(* IEC 61131-3 sources: Test-Git_ESME26/TestProgettoESME_26.fbsproj/AxisModuleLib Migration, 10 files *)

(* ---- AXM_GPL.gvl ---- *)
{attribute 'qualified_only'}
VAR_GLOBAL CONSTANT
	Gc_udiMaxNumberOfCamTables		: UDINT := 4;
END_VAR

(* ---- AXM_FC_EtCmdToString.fn.st ---- *)
FUNCTION PUBLIC AXM_FC_EtCmdToString : STRING[20]
VAR_INPUT
	i_etCmd : AXM_ET_Cmd;
END_VAR
VAR_OUTPUT
	q_etDiag	: GD.ET_Diag := GD.ET_Diag.Ok;
	q_etDiagExt	: AXM_ET_DiagExt := AXM_ET_DiagExt.Ok;
END_VAR
VAR
END_VAR

AXM_FC_EtCmdToString := TO_STRING(i_etCmd);
IF TO_UDINT(AXM_FC_EtCmdToString) <> 0 THEN // if the string is not a number the result is 0
	AXM_FC_EtCmdToString := Standard.CONCAT('Unknown DiagExt: ', TO_STRING(i_etCmd));
	q_etDiag := GD.ET_Diag.InputParameterInvalid;
	q_etDiagExt := AXM_ET_DiagExt.CmdUnknown;;
END_IF

(* ---- AXM_FC_EtMotionActiveVelTypeToString.fn.st ---- *)
FUNCTION PUBLIC AXM_FC_EtMotionActiveVelTypeToString : STRING[20]
VAR_INPUT
	i_etMotionActiveVelType : AXM_ET_MotionActiveVelType;
END_VAR
VAR_OUTPUT
	q_etDiag	: GD.ET_Diag := GD.ET_Diag.Ok;
	q_etDiagExt	: AXM_ET_DiagExt := AXM_ET_DiagExt.Ok;
END_VAR
VAR
END_VAR

AXM_FC_EtMotionActiveVelTypeToString := TO_STRING(i_etMotionActiveVelType);

(* ---- AXM_FC_EtOpModeToString.fn.st ---- *)
FUNCTION PUBLIC AXM_FC_EtOpModeToString : STRING[20]
VAR_INPUT
	i_etOpMode : AXM_ET_OpMode;
END_VAR
VAR_OUTPUT
	q_etDiag	: GD.ET_Diag := GD.ET_Diag.Ok;
	q_etDiagExt	: AXM_ET_DiagExt := AXM_ET_DiagExt.Ok;
END_VAR
VAR
END_VAR

AXM_FC_EtOpModeToString := TO_STRING(i_etOpMode);

(* ---- AXM_FC_EtParIdToString.fn.st ---- *)
FUNCTION PUBLIC AXM_FC_EtParIdToString : STRING[20]
VAR_INPUT
	i_etParId : AXM_ET_ParId;
END_VAR
VAR_OUTPUT
	q_etDiag	: GD.ET_Diag := GD.ET_Diag.Ok;
	q_etDiagExt	: AXM_ET_DiagExt := AXM_ET_DiagExt.Ok;
END_VAR
VAR
END_VAR

AXM_FC_EtParIdToString := TO_STRING(i_etParId);

(* ---- AXM_FC_EtStateToString.fn.st ---- *)
FUNCTION PUBLIC AXM_FC_EtStateToString : String[80]
VAR_INPUT
	i_etState	: AXM_ET_State;
END_VAR
VAR_OUTPUT
	q_etDiag	: GD.ET_Diag := GD.ET_Diag.Ok;
	q_etDiagExt	: AXM_ET_DiagExt := AXM_ET_DiagExt.Ok;
END_VAR
VAR
END_VAR

AXM_FC_EtStateToString := TO_STRING(i_etState);

(* ---- AXM_FC_UpdateAddInterfaceStruct.fn.st ---- *)
/// FC version: 1.0.0.0
/// Example Project version: 26.0.11.0 (Automatically generated, do not change!)

FUNCTION PUBLIC AXM_FC_UpdateAddInterfaceStruct : BOOL
VAR_INPUT
	i_pdwSubModuleAddInterfaces : POINTER TO TPL.TYPE_ADDRESS; // change from DWORD to TYPE_ADDRESS;
	i_udiSubModuleConstant		: UDINT;
END_VAR
VAR_IN_OUT
	iq_stAxisModuleItf	: AXM_ST_ModuleInterface;
END_VAR
VAR_OUTPUT
	q_etDiag			: GD.ET_Diag := GD.ET_Diag.Ok;
	q_etDiagExt			: AXM_ET_DiagExt := AXM_ET_DiagExt.Ok;
	q_sMsg				: STRING[80];
END_VAR
VAR
	pdwArrayPos			: POINTER TO TPL.TYPE_ADDRESS; // change from DWORD to TYPE_ADDRESS;
END_VAR

(********************************************************************************************************
revision history:
=========================================================================================================
version	|	date		| author				| comment
=========================================================================================================
1.0.0.0	|	2025-03-18	| Schneider Electric	| - initial release
---------------------------------------------------------------------------------------------------------
1.x.y.z	|	20xx-xx-xx	| your name				| - What has been modified?
=========================================================================================================
********************************************************************************************************)

IF i_pdwSubModuleAddInterfaces = 0 THEN
	q_etDiag	:= GD.ET_Diag.InputParameterInvalid;
	q_etDiagExt	:= AXM_ET_DiagExt.SubModuleAddInterfacesInvalidPointer;
	q_sMsg		:= '';
ELSIF i_udiSubModuleConstant < 1 THEN
	q_etDiag	:= GD.ET_Diag.InputParameterInvalid;
	q_etDiagExt := AXM_ET_DiagExt.SubModuleConstantRange;
	q_sMsg		:= '1 <= i_udiSubModuleConstant';
ELSE
	pdwArrayPos := i_pdwSubModuleAddInterfaces + (i_udiSubModuleConstant-1) * SIZEOF(pdwArrayPos^);
	pdwArrayPos^ := ADR(iq_stAxisModuleItf);
END_IF

(* ---- AXM_FB_AxisModuleController.fb.st ---- *)
FUNCTION_BLOCK PUBLIC AXM_FB_AxisModuleController
VAR_INPUT
	i_xEnable			: BOOL;
END_VAR
VAR_IN_OUT
	iq_stStandardModuleItf			: TPL.ST_StandardModuleInterface;
	iq_stStandardMotionItf			: TPL.ST_StandardMotionInterface;
	iq_stExceptionList				: TPL.ST_ExceptionList;
	iq_stLogDataList				: TPL.ST_LogDataList;
END_VAR
VAR_OUTPUT
	q_xActive			: BOOL;
	q_xReady			: BOOL;
	q_etDiag			: GD.ET_Diag := GD.ET_Diag.Ok;
	q_etDiagExt			: AXM_ET_DiagExt := AXM_ET_DiagExt.Disabled;
	q_sMsg				: STRING[80] := '';
END_VAR
VAR
	pdw								: POINTER TO TPL.TYPE_ADDRESS; // change from DWORD to TYPE_ADDRESS;
	udiModul						: UDINT;
	pstStandardInterface			: POINTER TO TPL.ST_StandardModuleInterface;
	pstAxisInterface				: POINTER TO AXM_ST_ModuleInterface;
	xSercState						: BOOL;
	xSercStateOld					: BOOL := TRUE;
	xJogForwEdgeDetect              : BOOL := FALSE;
	xJogBackEdgeDetect              : BOOL := FALSE;
END_VAR

IF i_xEnable AND NOT q_xActive THEN
	q_xActive := TRUE;
	q_xReady := TRUE;
	q_etDiag := GD.ET_Diag.Ok;
	q_etDiagExt := AXM_ET_DiagExt.Working;
	q_sMsg		:= '';
ELSIF NOT i_xEnable AND q_xActive THEN
	IF(iq_stStandardModuleItf.iq_stExt.dwSubModulesItf <> 0 AND iq_stStandardModuleItf.iq_stExt.pdwSubModulesAddItf <> 0) THEN
		FOR udiModul:= 1 TO iq_stStandardModuleItf.iq_stExt.udiNumberOfSubModules DO
			pstStandardInterface := iq_stStandardModuleItf.iq_stExt.dwSubModulesItf + UDINT_TO_DWORD((udiModul - 1) * SIZEOF(pstStandardInterface^));
			IF(pstStandardInterface^.q_dwModuleType = UDINT_TO_DWORD(TPL.ET_ModuleType.AxisModule)) THEN
				(* Module version check *)
				IF(pstStandardInterface^.q_udiModuleVersion = 1) THEN
					pdw := iq_stStandardModuleItf.iq_stExt.pdwSubModulesAddItf + UDINT_TO_DWORD((udiModul - 1) * SIZEOF(pdw^));
					pstAxisInterface := pdw^;
					IF(pstAxisInterface <> 0) THEN
						pstAxisInterface^.stManual.i_xJogForw := FALSE;
						pstAxisInterface^.stManual.i_xJogBack := FALSE;
					END_IF
				END_IF
			END_IF
		END_FOR
	END_IF
	q_xReady 	:= FALSE;
	q_xActive	:= FALSE;
	q_etDiag	:= GD.ET_Diag.Ok;
	q_etDiagExt	:= AXM_ET_DiagExt.Disabled;
	q_sMsg		:= '';
END_IF
IF ((iq_stStandardModuleItf.iq_stExt.udiNumberOfSubModules <> 0)
	AND ((iq_stStandardModuleItf.iq_stExt.pdwSubModulesAddItf = 0) OR (iq_stStandardModuleItf.iq_stExt.dwSubModulesItf = 0))) THEN
	q_xReady := FALSE;
	q_etDiag := GD.ET_Diag.InputParameterInvalid;
	q_etDiagExt := AXM_ET_DiagExt.MissingExtInit;
	q_sMsg := 'Missing Call of FC_UpdateAddInterfaceStruct';
END_IF

IF q_xActive AND q_xReady  THEN
 	IF (FC_GetSercosState() >= SMI.ET_SercosState.NRT) THEN
		xSercState := (FC_GetSercosState() = SMI.ET_SercosState.Phase4);
		IF(iq_stStandardModuleItf.iq_stExt.dwSubModulesItf <> 0 AND iq_stStandardModuleItf.iq_stExt.pdwSubModulesAddItf <> 0) THEN
			FOR udiModul := 1 TO iq_stStandardModuleItf.iq_stExt.udiNumberOfSubModules DO
				pstStandardInterface := iq_stStandardModuleItf.iq_stExt.dwSubModulesItf + UDINT_TO_DWORD((udiModul - 1) * SIZEOF(pstStandardInterface^));
				IF(pstStandardInterface^.q_dwModuleType = TPL.ET_ModuleType.AxisModule) THEN
					(* Module version check *)
					IF(pstStandardInterface^.q_udiModuleVersion = 1) THEN
						pdw := iq_stStandardModuleItf.iq_stExt.pdwSubModulesAddItf +  UDINT_TO_DWORD((udiModul - 1) * SIZEOF(pdw^));
						IF(pdw^ = 0) THEN (* Configuration error in stSubModules *)
							q_xReady := FALSE;
							q_etDiag := GD.ET_Diag.InputParameterInvalid;
							q_etDiagExt := AXM_ET_DiagExt.MissingExtInit;
							q_sMsg := 'Missing Call of FC_UpdateAddInterfaceStruct';
							RETURN;
						END_IF
						pstAxisInterface := pdw^;
						IF(pstAxisInterface <> 0) THEN
							(* Implementation of axis select *)
							IF iq_stStandardMotionItf.i_udiModuleSelect > 0 AND iq_stStandardMotionItf.i_udiModuleSelect = pstStandardInterface^.i_udiModuleId THEN

								(* Don't set pstAxisInterface^.stManual.i_xJog* from iq_stStandardMotionItf.i_xJog* blindly since the Vis might want to jog as well *)
								IF (iq_stStandardMotionItf.i_xJogForw) THEN
									pstAxisInterface^.stManual.i_xJogForw := TRUE;
									xJogForwEdgeDetect := TRUE;
								ELSE
									IF (xJogForwEdgeDetect) THEN
										pstAxisInterface^.stManual.i_xJogForw := FALSE;
										xJogForwEdgeDetect := FALSE;
								    END_IF
								END_IF
								IF (iq_stStandardMotionItf.i_xJogBack) THEN
									pstAxisInterface^.stManual.i_xJogBack := TRUE;
									xJogBackEdgeDetect := TRUE;
								ELSE
									IF (xJogBackEdgeDetect) THEN
										pstAxisInterface^.stManual.i_xJogBack := FALSE;
										xJogBackEdgeDetect := FALSE;
								    END_IF
								END_IF

							ELSE
								pstAxisInterface^.stManual.i_xJogForw := FALSE;
								pstAxisInterface^.stManual.i_xJogBack := FALSE;
							END_IF
							(* Implementation of HomeOkReset *)
							IF NOT xSercState  THEN (* As long as the sercos state is <> 4, set the reset home ok to true *)
								pstAxisInterface^.stHome.i_xResetHomeOk := TRUE;
							ELSIF NOT xSercStateOld THEN (* Detect a positive edge in xSercState, the sercos has entered state 4 *)
								pstAxisInterface^.stHome.i_xResetHomeOk := FALSE;
							END_IF
						END_IF
					END_IF
				END_IF
			END_FOR
 		END_IF
	ELSE
		xSercState := FALSE;
		q_xReady := FALSE;
		q_etDiag := GD.ET_Diag.SercosConditionInvalid;
		q_etDiagExt := AXM_ET_DiagExt.GlobalSercosInterfaceInvalid;
		q_sMsg := AXM_FC_EtDiagExtToString(i_etDiagExt := AXM_ET_DiagExt.GlobalSercosInterfaceInvalid);
	END_IF
	xSercStateOld := xSercState;
END_IF

(* ---- AXM_FB_AxisModuleVisController.fb.st ---- *)
FUNCTION_BLOCK PUBLIC AXM_FB_AxisModuleVisController
VAR_INPUT
	i_xEnable               : BOOL;
	i_pstMachineStandardItf : POINTER TO TPL.ST_StandardModuleInterface;
	i_pstCurrentStandardItf : POINTER TO TPL.ST_StandardModuleInterface;
	i_dwCurrentAddItf       : TPL.TYPE_ADDRESS; // change DWORD to TYPE_ADDRESS
	i_xUpdateData           : BOOL;
	i_udiCurrentJogTarget   : UDINT;
END_VAR
VAR_IN_OUT
	iq_stExceptionList : TPL.ST_ExceptionList;
	iq_stLogDataList   : TPL.ST_LogDataList;
END_VAR
VAR_OUTPUT
	q_xActive                          : BOOL;
	q_xReady                           : BOOL;
	q_etDiag                           : GD.ET_Diag := GD.ET_Diag.Ok;
	q_etDiagExt                        : AXM_ET_DiagExt := AXM_ET_DiagExt.Disabled;
	q_sMsg                             : STRING[80] := '';
	q_udiSetAsCurrentModule            : UDINT;
	q_udiSetAsJogTarget                : UDINT;
	q_xSimulateExceptionStopEndOfCycle : BOOL;
END_VAR
VAR
	xEnableFlag              : BOOL;
	pstCurrentAxisInterface  : POINTER TO AXM_ST_ModuleInterface;
	stOldAxisInterface       : AXM_ST_ModuleInterface;
	pstCurrent               : POINTER TO TPL.ST_StandardModuleInterface;
	xInitUserInputs          : BOOL;
	dwOldCurrentAddInterface : TPL.TYPE_ADDRESS; // change DWORD to TYPE_ADDRESS
	xSuccess                 : BOOL;
END_VAR
VAR
	viq_stCurrentAxisInterface      : AXM_ST_ModuleInterface;
	viq_pstCurrentStandardInterface : POINTER TO TPL.ST_StandardModuleInterface;
	vq_xCurrentIsOfMyType           : BOOL;
	vi_iPaneSelect                  : INT  := 1;
	vq_iShowOpMode                  : DINT := -1;
	vq_sOpMode                      : STRING[40];
	vi_iSelectOpMode                : INT  := -1;
	vq_sDriveName                   : STRING[40];
	vq_lrDriveRefPosition           : LREAL;
	vq_uiDriveTopologyAddress       : UINT;
	vq_diDriveState                 : DINT;
	vq_diDriveDiagCode              : DINT;
	vq_sDriveDiagMsg                : STRING[39];
	vq_lrDriveMaxVel                : LREAL;
	vq_lrDriveMaxAcc                : LREAL;
	vq_xDriveControllerEnable       : BOOL;
	vq_diDriveWorkingState          : DINT;
	vq_sMasterName                  : STRING[40];
	vq_xTpValue                     : BOOL;
	viq_xCmdStart                   : BOOL;
	viq_xCmdWSStart                 : BOOL;
	viq_xCmdHold                    : BOOL;
	viq_xDriveEnableOn              : BOOL;
	viq_xDriveEnableOff             : BOOL;
	viq_xReactionEndOfCycle         : BOOL;
	viq_xHomeLimitSwitchInvisible   : BOOL;
	viq_xHomeMoveOnPosInvisible     : BOOL;
	viq_xHomeSensorInvisible        : BOOL;
	viq_xHomeSetPosInvisible        : BOOL;
	viq_xHomeTorqueInvisible        : BOOL;
	viq_xHomeTouchProbeInvisible    : BOOL;
	viq_xHomeWritePosInvisible      : BOOL;
	viq_xHomeForceInvisible         : BOOL;
	viq_xJogForw                    : BOOL;
	viq_xJogBack                    : BOOL;
	xJogForwEdgeDetect              : BOOL := FALSE;
	xJogBackEdgeDetect              : BOOL := FALSE;
	viq_xEditCamTablesInvisible     : BOOL := TRUE;
	viq_udiEditCamTablesTableNo     : UDINT := 4;
	viq_diEditCamTablesPointNo      : DINT := 0;
	v_xHideTabHandler               : BOOL := TRUE;
	ifDiagnostic                    : UFMPLCI.IF_Diagnostic;
	ifDiagnosticAccess              : UFMPLCI.IF_DiagnosticAccess;
	ifGetParentDevice               : DTSI.IF_GetParentDevice;
	ifDeviceAccess                  : DTSI.IF_DeviceAccess;
	ifSercosIdentificationAccess    : SDI.IF_SercosIdentificationAccess;
	ifSercosIdentification          : SDI.IF_SercosIdentification;
	ifWorkingModeAccess             : CFDI.IF_WorkingModeAccess;
	ifWorkingMode                   : CFDI.IF_WorkingMode;
	ifDeviceTreeObjectSlaveAccess   : UFMPLCI.IF_DeviceTreeObjectAccess;
	ifDeviceTreeObjectMasterAccess  : UFMPLCI.IF_DeviceTreeObjectAccess;
	ifDriveConfigAccess             : DDI.IF_DriveConfigAccess;
	ifDriveConfig                   : DDI.IF_DriveConfig;
	ifOldMaster                     : MOIN.IF_Axis;
	ifTouprobeData                  : IODI.IF_TouchprobeData;
	ifTouprobeDataAccess            : IODI.IF_TouchprobeDataAccess;

END_VAR

q_udiSetAsCurrentModule            := 0;
q_udiSetAsJogTarget                := 0;
pstCurrent                         := i_pstCurrentStandardItf;
q_xSimulateExceptionStopEndOfCycle := viq_xReactionEndOfCycle;

// Calculate Homing mode invisible BOOLs
viq_xHomeLimitSwitchInvisible := viq_stCurrentAxisInterface.stHome.i_etMode < 8 OR viq_stCurrentAxisInterface.stHome.i_etMode > 11;
viq_xHomeMoveOnPosInvisible   := viq_stCurrentAxisInterface.stHome.i_etMode <> 14;
viq_xHomeSensorInvisible      := viq_stCurrentAxisInterface.stHome.i_etMode < 4 OR viq_stCurrentAxisInterface.stHome.i_etMode > 7;
viq_xHomeSetPosInvisible      := viq_stCurrentAxisInterface.stHome.i_etMode < 15 OR viq_stCurrentAxisInterface.stHome.i_etMode > 19;
viq_xHomeTorqueInvisible      := viq_stCurrentAxisInterface.stHome.i_etMode < 12 OR viq_stCurrentAxisInterface.stHome.i_etMode > 13;
viq_xHomeTouchProbeInvisible  := viq_stCurrentAxisInterface.stHome.i_etMode < 0 OR viq_stCurrentAxisInterface.stHome.i_etMode > 3;
viq_xHomeWritePosInvisible    := viq_stCurrentAxisInterface.stHome.i_etMode <> 20;
viq_xHomeForceInvisible       := viq_stCurrentAxisInterface.stHome.i_etMode < 21 OR viq_stCurrentAxisInterface.stHome.i_etMode > 22;

IF i_xEnable THEN
	q_xActive := TRUE;
	IF (i_pstCurrentStandardItf = 0) THEN
		q_xReady    := FALSE;
		q_etDiag    := GD.ET_Diag.InputParameterInvalid;
		q_etDiagExt := AXM_ET_DiagExt.CurrentStandardItfInvalid;
		q_sMsg      := 'pointer is null';
	ELSIF (i_dwCurrentAddItf = 0) THEN
		q_xReady    := FALSE;
		q_etDiag    := GD.ET_Diag.InputParameterInvalid;
		q_etDiagExt := AXM_ET_DiagExt.CurrentAddItfInvalid;
		q_sMsg      := 'pointer is null';
	ELSE
		q_xReady    := TRUE;
		q_etDiag    := GD.ET_Diag.Ok;
		q_etDiagExt := AXM_ET_DiagExt.Working;
		q_sMsg      := AXM_FC_EtDiagExtToString(i_etDiagExt := AXM_ET_DiagExt.Working);
		IF (i_pstCurrentStandardItf^.q_dwModuleType = UDINT_TO_DWORD(TPL.ET_ModuleType.AxisModule)) THEN
			(* Module version check *)
			IF (i_pstCurrentStandardItf^.q_udiModuleVersion = 1) THEN
				pstCurrentAxisInterface := i_dwCurrentAddItf;
				vq_xCurrentIsOfMyType   := TRUE;
			END_IF
		ELSE
			pstCurrentAxisInterface := 0;
			vq_xCurrentIsOfMyType   := FALSE;
		END_IF

		IF (vq_xCurrentIsOfMyType) THEN
			(* Execute changes requested by user first *)
			IF (NOT xInitUserInputs) THEN
				xInitUserInputs := TRUE;
				(* Ignore values of variables now *)
			ELSE
				DetectUserChanges();
			END_IF

			IF dwOldCurrentAddInterface <> i_dwCurrentAddItf THEN
				dwOldCurrentAddInterface        := i_dwCurrentAddItf;
				viq_stCurrentAxisInterface      := pstCurrentAxisInterface^;
				stOldAxisInterface              := viq_stCurrentAxisInterface;
				viq_pstCurrentStandardInterface := i_pstCurrentStandardItf;

				IF (viq_stCurrentAxisInterface.stMain.i_ifDrive <> 0) THEN
					xSuccess := __QUERYINTERFACE(viq_stCurrentAxisInterface.stMain.i_ifDrive, ifGetParentDevice);
					IF xSuccess THEN
						ifDeviceAccess := ifGetParentDevice.GetParentDevice();
						xSuccess       := __QUERYINTERFACE(ifDeviceAccess, ifDiagnosticAccess);
						IF xSuccess THEN
							ifDiagnostic := ifDiagnosticAccess.Diagnostic;
						END_IF
						xSuccess := __QUERYINTERFACE(ifDeviceAccess, ifDriveConfigAccess);
						IF xSuccess THEN
							ifDriveConfig := ifDriveConfigAccess.DriveConfig;
						END_IF
						xSuccess := __QUERYINTERFACE(ifDeviceAccess, ifDeviceTreeObjectSlaveAccess);
						IF xSuccess THEN
							vq_sDriveName := ifDeviceTreeObjectSlaveAccess.DeviceTreeObject.Name;
						END_IF
						xSuccess := __QUERYINTERFACE(ifDeviceAccess, ifSercosIdentificationAccess);
						IF xSuccess THEN
							ifSercosIdentification := ifSercosIdentificationAccess.SercosIdentification;
						END_IF
						xSuccess := __QUERYINTERFACE(ifDeviceAccess, ifWorkingModeAccess);
						IF xSuccess THEN
							ifWorkingMode := ifWorkingModeAccess.WorkingMode;
						END_IF
					ELSE
						vq_sDriveName := '';
					END_IF
				END_IF
				IF viq_stCurrentAxisInterface.stHome.stTouchProbe.i_ifTouchProbe <> 0 THEN
					xSuccess := __QUERYINTERFACE(viq_stCurrentAxisInterface.stHome.stTouchProbe.i_ifTouchProbe, ifGetParentDevice);
					IF xSuccess THEN
						ifDeviceAccess := ifGetParentDevice.GetParentDevice();
						xSuccess       := __QUERYINTERFACE(ifDeviceAccess, ifTouprobeDataAccess);
						IF xSuccess THEN
							ifTouprobeData := ifTouprobeDataAccess.TouchprobeData;
						END_IF
					END_IF
				END_IF
			END_IF

			(* generate VisData *)
			IF (vi_iSelectOpMode < 0) THEN
				(* Show actual OpMode *)
				vq_ishowOpMode := DINT_TO_INT(viq_stCurrentAxisInterface.stMain.q_etOpMode);
			ELSE
				vq_ishowOpMode := vi_iSelectOpMode;
			END_IF

			IF (viq_stCurrentAxisInterface.stMain.i_ifDrive <> 0) THEN
				vq_diDriveState       := TO_DINT(viq_stCurrentAxisInterface.stMain.i_ifDrive.etAxisState);
				vq_lrDriveRefPosition := viq_stCurrentAxisInterface.stMain.i_ifDrive.lrPosition;
				vq_sOpMode            := AXM_FC_EtOpModeToString(i_etOpMode := viq_stCurrentAxisInterface.stMain.q_etOpMode);
			END_IF

			IF ifDiagnostic <> 0 THEN
				vq_diDriveDiagCode := ifDiagnostic.DiagCode;
				vq_sDriveDiagMsg   := ifDiagnostic.DiagMsg;
			ELSE
				vq_diDriveDiagCode := 0;
				vq_sDriveDiagMsg   := '';
			END_IF

			IF ifSercosIdentification <> 0 THEN
				vq_uiDriveTopologyAddress := ifSercosIdentification.TopologyAddress;
			ELSE
				vq_uiDriveTopologyAddress := 0;
			END_IF

			IF ifWorkingMode <> 0 THEN
				vq_diDriveWorkingState := ifWorkingMode.ActualState;
			ELSE
				vq_diDriveWorkingState := 0;
			END_IF

			IF (viq_stCurrentAxisInterface.stMain.i_ifDrive <> 0) THEN
				vq_lrDriveRefPosition := viq_stCurrentAxisInterface.stMain.i_ifDrive.lrPosition;
				vq_sOpMode            := AXM_FC_EtOpModeToString(i_etOpMode := viq_stCurrentAxisInterface.stMain.q_etOpMode);

				IF ifDriveConfig = 0 THEN
					vq_lrDriveMaxVel := 0.0;
					vq_lrDriveMaxAcc := 0.0;
				ELSE
					vq_lrDriveMaxVel := ifDriveConfig.MaxVel;
					vq_lrDriveMaxAcc := ifDriveConfig.MaxAcc;
				END_IF

				//xSuccess := __QUERYINTERFACE(viq_stCurrentAxisInterface.stMain.i_ifDrive, ifDrivePowerControlMandatory);
				//IF NOT xSuccess OR (ifDrivePowerControlMandatory = 0) THEN
				//	(* ignore error *)
				//	ifDrivePowerControlMandatory := 0;
				//	vq_xDriveControllerEnable := FALSE;
				//ELSE
				//	vq_xDriveControllerEnable := ifDrivePowerControlMandatory.ControllerEnable;
				//END_IF
			ELSE
				vq_xDriveControllerEnable := FALSE;
				vq_lrDriveMaxVel          := 0.0;
				vq_lrDriveMaxAcc          := 0.0;
				vq_lrDriveRefPosition     := 0.0;
			END_IF

			IF (viq_stCurrentAxisInterface.stMain.i_ifMaster <> 0) THEN
				IF ifOldMaster <> viq_stCurrentAxisInterface.stMain.i_ifMaster THEN
					ifOldMaster := viq_stCurrentAxisInterface.stMain.i_ifMaster;
					xSuccess    := __QUERYINTERFACE(viq_stCurrentAxisInterface.stMain.i_ifMaster, ifGetParentDevice);
					IF xSuccess THEN
						ifDeviceAccess := ifGetParentDevice.GetParentDevice();
						xSuccess       := __QUERYINTERFACE(ifDeviceAccess, ifDeviceTreeObjectMasterAccess);
						IF xSuccess THEN
							vq_sMasterName := ifDeviceTreeObjectMasterAccess.DeviceTreeObject.Name;
						END_IF
					ELSE
						//no device tree object
						vq_sMasterName := '';
					END_IF
				END_IF
			ELSE
				vq_sMasterName := 'not set';
			END_IF

			IF (ifTouprobeData <> 0) THEN
				vq_xTpValue := ifTouprobeData.Value;
			ELSE
				vq_xTpValue := FALSE;
			END_IF

			IF iq_stExceptionList.udiNumberOfActiveExceptions > 0 AND viq_stCurrentAxisInterface.stMain.q_etOpMode = AXM_ET_OpMode.NoOp THEN
				pstCurrentAxisInterface^.stMain.i_xStart   := FALSE;
				viq_stCurrentAxisInterface.stMain.i_xStart := FALSE;
				stOldAxisInterface.stMain.i_xStart         := FALSE;

				pstCurrentAxisInterface^.stPos.i_xStop   := FALSE;
				viq_stCurrentAxisInterface.stPos.i_xStop := FALSE;
				stOldAxisInterface.stPos.i_xStop         := FALSE;
			END_IF

			IF (viq_xJogForw) THEN
				viq_stCurrentAxisInterface.stManual.i_xJogForw := TRUE;
				xJogForwEdgeDetect                             := TRUE;
			ELSE
				IF (xJogForwEdgeDetect) THEN
					viq_stCurrentAxisInterface.stManual.i_xJogForw := FALSE;
					xJogForwEdgeDetect                             := FALSE;
				END_IF
			END_IF

			IF (viq_xJogBack) THEN
				viq_stCurrentAxisInterface.stManual.i_xJogBack := TRUE;
				xJogBackEdgeDetect                             := TRUE;
			ELSE
				IF (xJogBackEdgeDetect) THEN
					viq_stCurrentAxisInterface.stManual.i_xJogBack := FALSE;
					xJogBackEdgeDetect                             := FALSE;
				END_IF
			END_IF

			IF (i_udiCurrentJogTarget <> i_pstCurrentStandardItf^.i_udiModuleId) AND (viq_xJogForw OR viq_xJogBack) THEN
				q_udiSetAsJogTarget                            := i_pstCurrentStandardItf^.i_udiModuleId; (* select as jog target whenever a jog button is pushed *)
				viq_stCurrentAxisInterface.stManual.i_xJogForw := FALSE;
				viq_stCurrentAxisInterface.stManual.i_xJogBack := FALSE;
			END_IF

		ELSE
			;
		END_IF
	END_IF
ELSE
	vq_xCurrentIsOfMyType := FALSE;
	q_xActive             := FALSE;
	q_xReady              := FALSE;
	q_etDiag              := GD.ET_Diag.Ok;
	q_etDiagExt           := AXM_ET_DiagExt.Disabled;
	q_sMsg                := AXM_FC_EtDiagExtToString(i_etDiagExt := AXM_ET_DiagExt.Disabled);
END_IF

(* ---- AXM_FB_TabSwitch.fb.st ---- *)
FUNCTION_BLOCK AXM_FB_TabSwitch
VAR_INPUT
	i_xEnable				: BOOL;
	i_xLowEnd				: BOOL;
	i_xHighEnd				: BOOL;
	i_udiTableSelectNr		: UDINT;
END_VAR
VAR_IN_OUT
	iq_xTakeNewCam			: BOOL;
	iq_xTakeInstantNewCam	: BOOL;
	iq_xNewCam				: BOOL;
	iq_xInstantNewCam		: BOOL;
	iq_astMotionPar			: ARRAY [0..AXM_GPL.Gc_udiMaxNumberOfCamTables] OF CMT.ST_MultiCam;
	iq_stOutTab				: CMT.ST_MultiCam;
END_VAR
VAR_OUTPUT
	q_xActive				: BOOL;
	q_xReady				: BOOL;
	q_etDiag				: GD.ET_Diag := GD.ET_Diag.Ok;
	q_etDiagExt				: AXM_ET_DiagExt := AXM_ET_DiagExt.Disabled;
	q_sMsg					: STRING[80] := '';
	q_udiTableNumber		: UDINT;
END_VAR
VAR
	xEnableFlag				: BOOL;
	diState					: DINT;
	udiTableSelectNr_old	: UDINT := AXM_GPL.Gc_udiMaxNumberOfCamTables +1;
	xWaitNewCamAccept		: BOOL;
END_VAR

IF i_xEnable AND NOT xEnableFlag AND (diState = 0) THEN
	xEnableFlag := TRUE;
	q_xActive := TRUE;
	q_xReady := TRUE;
	q_etDiag := GD.ET_Diag.Ok;
	q_etDiagExt := AXM_ET_DiagExt.Working;
	q_sMsg := AXM_FC_EtDiagExtToString(i_etDiagExt := AXM_ET_DiagExt.Working);
	iq_xTakeNewCam := FALSE;
	iq_xTakeInstantNewCam := FALSE;
	iq_xNewCam := FALSE;
	iq_xInstantNewCam := FALSE;
	IF (i_udiTableSelectNr <= AXM_GPL.Gc_udiMaxNumberOfCamTables) THEN
		iq_stOutTab := iq_astMotionPar[i_udiTableSelectNr];
		q_udiTableNumber := i_udiTableSelectNr;
		IF udiTableSelectNr_old = AXM_GPL.Gc_udiMaxNumberOfCamTables +1 THEN
			// on very first call after controller boot FB_MultiCam has not seen any new cam, therefore set of iq_xNewCam in state 10 would cause that a non cyclic cam is executed twice
			udiTableSelectNr_old := i_udiTableSelectNr;
		END_IF
	ELSE
		iq_stOutTab := iq_astMotionPar[0];
		q_udiTableNumber := 0;
	END_IF
	//udiTableSelectNr_old := i_udiTableSelectNr;
	IF(xWaitNewCamAccept) THEN
		(* we did send a newcam, but the multicam has been disabled bevore he did compute it
			and beeing activated (or inactive) he resets the newcam so the signal is lost,
			but we do keep track ==> send it again *)
		diState := 1; (* special startup state *)
	ELSE
		diState:=10;
	END_IF
ELSIF NOT i_xEnable AND xEnableFlag THEN
	xEnableFlag := FALSE;
	q_xReady := FALSE;
	q_xActive := FALSE;
	q_etDiag := GD.ET_Diag.Ok;
	q_etDiagExt := AXM_ET_DiagExt.Disabled;
	q_sMsg := AXM_FC_EtDiagExtToString(i_etDiagExt := AXM_ET_DiagExt.Disabled);
	diState := 0;
END_IF

CASE diState OF
	0: (* Disabled *)
		; (* Do nothing *)

	1:
		(* send xNewCam in seccond cycle, because multicam does set iq_xNewCam to false when he is enabled *)
		iq_xNewCam := TRUE; (* if the fb was disabled before the multicam did compute the newcam,
			send a newCam signal to the multicam one cycle after he has been activated *)
		diState := 10;

	10: (* working *)
		IF iq_xTakeInstantNewCam THEN
			IF (i_udiTableSelectNr <= AXM_GPL.Gc_udiMaxNumberOfCamTables) THEN
				iq_stOutTab := iq_astMotionPar[i_udiTableSelectNr];
				q_udiTableNumber := i_udiTableSelectNr;
				udiTableSelectNr_old := i_udiTableSelectNr;
			ELSE
				iq_stOutTab := iq_astMotionPar[0];
				q_udiTableNumber := 0;
				udiTableSelectNr_old := 0;
			END_IF
			iq_xInstantNewCam := TRUE;
			diState := 30;
		ELSIF (i_xLowEnd OR i_xHighEnd) AND iq_xNewCam THEN
			diState :=20;
			iq_xTakeNewCam:= FALSE;
		ELSIF ((i_udiTableSelectNr <> udiTableSelectNr_old) OR iq_xTakeNewCam) AND NOT i_xLowEnd AND NOT i_xHighEnd THEN
			IF (i_udiTableSelectNr <= AXM_GPL.Gc_udiMaxNumberOfCamTables) THEN
				iq_stOutTab := iq_astMotionPar[i_udiTableSelectNr];
				q_udiTableNumber := i_udiTableSelectNr;
				udiTableSelectNr_old := i_udiTableSelectNr;
			ELSE
				iq_stOutTab := iq_astMotionPar[0];
				q_udiTableNumber := 0;
				udiTableSelectNr_old := 0;
			END_IF
			iq_xNewCam := TRUE;
			xWaitNewCamAccept := TRUE;
		END_IF
		IF (NOT iq_xNewCam) THEN
			xWaitNewCamAccept := FALSE;
		END_IF

	20: (* wait new cam accept *)
		IF NOT i_xLowEnd AND NOT i_xHighEnd  THEN
			diState:=10;
		END_IF
		IF(NOT iq_xNewCam) THEN
			xWaitNewCamAccept := FALSE;
		END_IF

	30: (* wait InstantNewCam accepted *)
		IF NOT iq_xInstantNewCam THEN
			iq_xTakeInstantNewCam := FALSE;
			diState := 10;
		END_IF
END_CASE
